Fanuc KAREL source: kb00052.KL

-- PROVISIONAL review KL for V1013-1; original PC SHA256 ef1e2aa41c39af628bbc2841c6ad96067ee8620d4f6f772102f57486c8d9d4ef
-- Incomplete behavior may be omitted. Consult companion uncertainty JSON. Do not deploy.
PROGRAM KB00052
%NOLOCKGROUP
VAR
  P1 : INTEGER
  P2 : INTEGER
-- UNRESOLVED_DECL RESULT type=000106
BEGIN
  -- UNRESOLVED_PC offsets 5-12; opcodes 9D,23
  -- UNRESOLVED_PC offsets 17-24; opcodes 9D,23
  -- UNRESOLVED_PC offsets 29-58; opcodes 27,22,22,27,9D,76,7E,4A
  -- UNRESOLVED_PC offsets 63-67; opcodes 7F
END KB00052
